{attribute 'qualified_only'}
{attribute 'strict'}
{attribute 'to_string'}
TYPE E_Line_Target :
(
	eNone := 0,
	eClose,
	eTank_A,
	eTank_B,
	eCIP,
	eDrain
);
END_TYPE

(* stored: Version 1.1.0.1, ProductVersion 3.1.4024.12
   EnumerationTextList E_Line_Target: Id {78a70d41-3ccd-4ccb-a601-f262cf1739ee} *)
